TYPE "ST_PressDemoUnitHal"
VERSION : 0.1
   STRUCT
      PressRam { ExternalAccessible := 'False'; ExternalVisible := 'False'; ExternalWritable := 'False'} : "ST_CylinderHal";
      Door { ExternalAccessible := 'False'; ExternalVisible := 'False'; ExternalWritable := 'False'} : "ST_CylinderHal";
      PartSlide { ExternalAccessible := 'False'; ExternalVisible := 'False'; ExternalWritable := 'False'} : "ST_CylinderHal";
   END_STRUCT;

END_TYPE

